(* IEC 61131-3 sources: model-first-plc-agent-ai/results/T1-W-27, 2 files *)

(* ---- a1_code.st ---- *)
FUNCTION_BLOCK ConveyorRuntime
VAR_INPUT
    sensor_a : BOOL;
    sensor_b : BOOL;
END_VAR
VAR_OUTPUT
    conveyor : BOOL := FALSE;
END_VAR
VAR
    command_latch : RS;
    x0 : BOOL := TRUE;
    x1 : BOOL := FALSE;
END_VAR

command_latch(
    S := sensor_a AND NOT sensor_b,
    R1 := sensor_b
);

x1 := command_latch.Q1;
x0 := NOT x1;
conveyor := x1;

END_FUNCTION_BLOCK

PROGRAM Main
VAR
    SensorA AT %IX100.0 : BOOL;
    SensorB AT %IX100.1 : BOOL;
    Conveyor AT %QX100.0 : BOOL;
END_VAR
VAR
    runtime : ConveyorRuntime;
    initialized : BOOL := FALSE;
END_VAR

IF NOT initialized THEN
    Conveyor := FALSE;
    initialized := TRUE;
END_IF;

runtime(
    sensor_a := SensorA,
    sensor_b := SensorB
);

Conveyor := runtime.conveyor;

END_PROGRAM

(* ---- a2_code.st ---- *)
FUNCTION_BLOCK FB_TransferControl
VAR_INPUT
    sensor_a : BOOL;
    sensor_b : BOOL;
END_VAR
VAR_OUTPUT
    conveyor : BOOL;
END_VAR
VAR
    conveyor_latch : RS;
END_VAR

conveyor_latch(
    S := sensor_a AND NOT sensor_b,
    R1 := sensor_b
);
conveyor := conveyor_latch.Q1;

END_FUNCTION_BLOCK

PROGRAM Main
VAR
    sensor_a AT %IX100.0 : BOOL;
    sensor_b AT %IX100.1 : BOOL;
    conveyor AT %QX100.0 : BOOL;
END_VAR
VAR
    transfer_control : FB_TransferControl;
END_VAR

transfer_control(
    sensor_a := sensor_a,
    sensor_b := sensor_b
);
conveyor := transfer_control.conveyor;

END_PROGRAM
